TYPE ST_PersistentRecipe :
STRUCT
	stInner : ST_PersistentInner;
	eMode : E_FixtureMode;
	sName : STRING(20);
	wsName : WSTRING(20);
	tDelay : TIME := T#1S500MS;
	dtStamp : DT;
	aPos : ARRAY[1..5] OF LREAL;
END_STRUCT
END_TYPE

(* stored: Version 1.1.0.1
   DUT ST_PersistentRecipe: Id {3f6a1c52-8d7e-4b0a-9a41-5c2e7d9b1a02} *)
